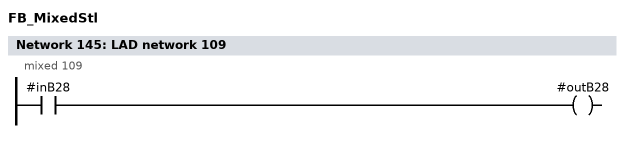
   RUNG wire#powerrail
      Contact( #inB28 )
      Coil( #outB28 )
   END_RUNG
   // the same network as SCL:
   #outB28 := #inB28;
END_REGION

REGION Network 146 (FBD): FBD network 110
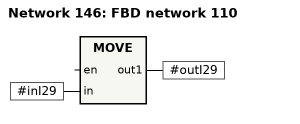
   #outI29 := #inI29;
END_REGION

REGION Network 147 (SCL): SCL network 111
   #tI10 := #inI30 + #cI20;
           IF #inB30 THEN
               #outR10 := #inR10 * 2.0;
           END_IF;
END_REGION

REGION Network 148 (STL): STL network 37
         A     #inB36;
         AN    #stB36;
         =     #outB36;
END_REGION

REGION Network 149: LAD network 112
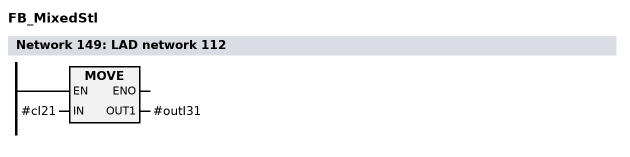
   RUNG wire#powerrail
      Move(in := #cI21, out1 => #outI31)
   END_RUNG
   // the same network as SCL:
   #outI31 := #cI21;
END_REGION

REGION Network 150 (FBD): FBD network 113
   // mixed 113
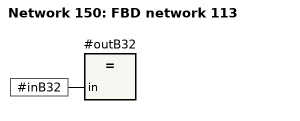
   #outB32 := #inB32;
END_REGION

REGION Network 151 (SCL): SCL network 114
   #tI13 := #inI33 + #cI23;
           IF #inB33 THEN
               #outR13 := #inR13 * 2.0;
           END_IF;
END_REGION

REGION Network 152 (STL): STL network 38
         L     #inI37;
         L     #stI37;
         +I;
         T     #outI37;
END_REGION

REGION Network 153: LAD network 115
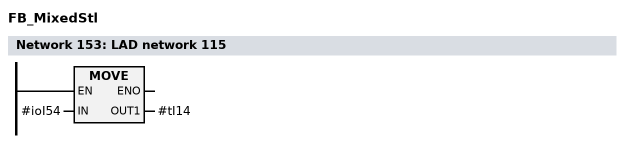
   RUNG wire#powerrail
      Move(in := #ioI54, out1 => #tI14)
   END_RUNG
   // the same network as SCL:
   #tI14 := #ioI54;
END_REGION

REGION Network 154 (FBD): FBD network 116
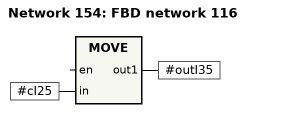
   #outI35 := #cI25;
END_REGION

REGION Network 155 (SCL): SCL network 117
   // mixed 117
   #tI16 := #inI36 + #cI26;
           IF #inB36 THEN
               #outR16 := #inR16 * 2.0;
           END_IF;
END_REGION

REGION Network 156 (STL): STL network 39
         L     #inR18;
         L     #tR38;
         *R;
         T     #outR18;  // product
END_REGION

REGION Network 157: LAD network 118
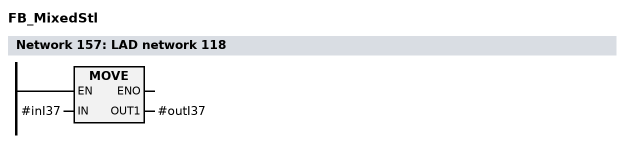
   RUNG wire#powerrail
      Move(in := #inI37, out1 => #outI37)
   END_RUNG
   // the same network as SCL:
   #outI37 := #inI37;
END_REGION

REGION Network 158 (FBD): FBD network 119
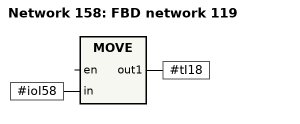
   #tI18 := #ioI58;
END_REGION

REGION Network 159 (SCL): SCL network 120
   #tI19 := #inI39 + #cI29;
           IF #inB39 THEN
               #outR19 := #inR19 * 2.0;
           END_IF;
END_REGION

REGION Network 160 (STL): STL network 40
         A     #inB39;
         AN    #stB39;
         =     #outB39;
END_REGION
END_FUNCTION_BLOCK

FUNCTION "FC_Stl" : Void   // FC1, STL
TITLE = STL test FC
{ S7_Optimized_Access := 'TRUE' }
VERSION : 0.1
   VAR_INPUT
      "a" : Bool;
      "b" : Bool;
      x : Int;
      y : Int;
   END_VAR
   VAR_OUTPUT
      q : Bool;
      sum : Int;
   END_VAR
   VAR_TEMP
      t : Int;
   END_VAR
BEGIN

REGION Network 1: Bit logic
   // Network comment line 1
         A     #"a";  // and a
         AN    #"b";
         =     #q;
END_REGION

REGION Network 2: Arithmetic
         L     #x;
         L     #y;
         +I;
         T     #t;

         L     #t;
         L     0;
         >I;
         JC    M001;
         L     0;
         T     #t;
   M001: L     #t;
         T     #sum;
END_REGION
END_FUNCTION

FUNCTION "FC_StlNoPar" : Void   // FC2, STL
{ S7_Optimized_Access := 'FALSE' }
VERSION : 0.1
BEGIN

REGION Network 1
         NOP   0;
END_REGION
END_FUNCTION

FUNCTION "FC_StlPar" : Void   // FC3, STL
{ S7_Optimized_Access := 'TRUE' }
VERSION : 0.1
   VAR_INPUT
      x : Int;
      y : Int;
   END_VAR
   VAR_OUTPUT
      q : Bool;
      r : Int;
   END_VAR
BEGIN

REGION Network 1
         L     #x;
         L     #y;
         +I;
         T     #r;
         >I;
         =     #q;
END_REGION
END_FUNCTION

FUNCTION "FC_BigFbd" : Void   // FC4, FBD
{ S7_Optimized_Access := 'TRUE' }
VERSION : 0.1
   VAR_INPUT
      inB0 : Bool;   // input bit 0
      inB1 : Bool;
      inB2 : Bool;
      inB3 : Bool;
      inB4 : Bool;
      inB5 : Bool;
      inB6 : Bool;
      inB7 : Bool;
      inB8 : Bool;
      inB9 : Bool;
      inB10 : Bool;   // input bit 10
      inB11 : Bool;
      inB12 : Bool;
      inB13 : Bool;
      inB14 : Bool;
      inB15 : Bool;
      inB16 : Bool;
      inB17 : Bool;
      inB18 : Bool;
      inB19 : Bool;
      inI0 : Int;
      inI1 : Int;
      inI2 : Int;
      inI3 : Int;
      inI4 : Int;
      inI5 : Int;
      inI6 : Int;
      inI7 : Int;
      inI8 : Int;
      inI9 : Int;
      inI10 : Int;
      inI11 : Int;
      inI12 : Int;
      inI13 : Int;
      inI14 : Int;
      inI15 : Int;
      inI16 : Int;
      inI17 : Int;
      inI18 : Int;
      inI19 : Int;
      inR0 : Real;
      inR1 : Real;
      inR2 : Real;
      inR3 : Real;
      inR4 : Real;
      inR5 : Real;
      inR6 : Real;
      inR7 : Real;
      inR8 : Real;
      inR9 : Real;
      inD0 : DInt;
      inD1 : DInt;
      inD2 : DInt;
      inD3 : DInt;
      inD4 : DInt;
      inD5 : DInt;
      inD6 : DInt;
      inD7 : DInt;
      inD8 : DInt;
      inD9 : DInt;
      inArr : Array[0..99] of Int;   // input array
      inStr : String;
      inSt : Struct
         x : Int;
         y : Real;
         z : Bool;
      END_STRUCT;
   END_VAR
   VAR_OUTPUT
      outB0 : Bool;
      outB1 : Bool;
      outB2 : Bool;
      outB3 : Bool;
      outB4 : Bool;
      outB5 : Bool;
      outB6 : Bool;
      outB7 : Bool;
      outB8 : Bool;
      outB9 : Bool;
      outB10 : Bool;
      outB11 : Bool;
      outB12 : Bool;
      outB13 : Bool;
      outB14 : Bool;
      outB15 : Bool;
      outB16 : Bool;
      outB17 : Bool;
      outB18 : Bool;
      outB19 : Bool;
      outI0 : Int;   // output int 0
      outI1 : Int;
      outI2 : Int;
      outI3 : Int;
      outI4 : Int;
      outI5 : Int;
      outI6 : Int;
      outI7 : Int;
      outI8 : Int;
      outI9 : Int;
      outI10 : Int;   // output int 10
      outI11 : Int;
      outI12 : Int;
      outI13 : Int;
      outI14 : Int;
      outI15 : Int;
      outI16 : Int;
      outI17 : Int;
      outI18 : Int;
      outI19 : Int;
      outR0 : Real;
      outR1 : Real;
      outR2 : Real;
      outR3 : Real;
      outR4 : Real;
      outR5 : Real;
      outR6 : Real;
      outR7 : Real;
      outR8 : Real;
      outR9 : Real;
      outD0 : DInt;
      outD1 : DInt;
      outD2 : DInt;
      outD3 : DInt;
      outD4 : DInt;
      outD5 : DInt;
      outD6 : DInt;
      outD7 : DInt;
      outD8 : DInt;
      outD9 : DInt;
   END_VAR
   VAR_IN_OUT
      ioI0 : Int;
      ioI1 : Int;
   END_VAR
   VAR_TEMP
      tI0 : Int;
      tI1 : Int;
      tI2 : Int;
      tI3 : Int;
      tI4 : Int;
      tI5 : Int;
      tI6 : Int;
      tI7 : Int;
      tI8 : Int;
      tI9 : Int;
      tI10 : Int;
      tI11 : Int;
      tI12 : Int;
      tI13 : Int;
      tI14 : Int;
      tI15 : Int;
      tI16 : Int;
      tI17 : Int;
      tI18 : Int;
      tI19 : Int;
      tI20 : Int;
      tI21 : Int;
      tI22 : Int;
      tI23 : Int;
      tI24 : Int;
      tI25 : Int;
      tI26 : Int;
      tI27 : Int;
      tI28 : Int;
      tI29 : Int;
      tI30 : Int;
      tI31 : Int;
      tI32 : Int;
      tI33 : Int;
      tI34 : Int;
      tI35 : Int;
      tI36 : Int;
      tI37 : Int;
      tI38 : Int;
      tI39 : Int;
      tI40 : Int;
      tI41 : Int;
      tI42 : Int;
      tI43 : Int;
      tI44 : Int;
      tI45 : Int;
      tI46 : Int;
      tI47 : Int;
      tI48 : Int;
      tI49 : Int;
      tI50 : Int;
      tI51 : Int;
      tI52 : Int;
      tI53 : Int;
      tI54 : Int;
      tI55 : Int;
      tI56 : Int;
      tI57 : Int;
      tI58 : Int;
      tI59 : Int;
      tI60 : Int;
      tI61 : Int;
      tI62 : Int;
      tI63 : Int;
      tI64 : Int;
      tI65 : Int;
      tI66 : Int;
      tI67 : Int;
      tI68 : Int;
      tI69 : Int;
      tI70 : Int;
      tI71 : Int;
      tI72 : Int;
      tI73 : Int;
      tI74 : Int;
      tI75 : Int;
      tI76 : Int;
      tI77 : Int;
      tI78 : Int;
      tI79 : Int;
      tI80 : Int;
      tI81 : Int;
      tI82 : Int;
      tI83 : Int;
      tI84 : Int;
      tI85 : Int;
      tI86 : Int;
      tI87 : Int;
      tI88 : Int;
      tI89 : Int;
      tI90 : Int;
      tI91 : Int;
      tI92 : Int;
      tI93 : Int;
      tI94 : Int;
      tI95 : Int;
      tI96 : Int;
      tI97 : Int;
      tI98 : Int;
      tI99 : Int;
      tR0 : Real;
      tR1 : Real;
      tR2 : Real;
      tR3 : Real;
      tR4 : Real;
      tR5 : Real;
      tR6 : Real;
      tR7 : Real;
      tR8 : Real;
      tR9 : Real;
      tR10 : Real;
      tR11 : Real;
      tR12 : Real;
      tR13 : Real;
      tR14 : Real;
      tR15 : Real;
      tR16 : Real;
      tR17 : Real;
      tR18 : Real;
      tR19 : Real;
      tR20 : Real;
      tR21 : Real;
      tR22 : Real;
      tR23 : Real;
      tR24 : Real;
      tR25 : Real;
      tR26 : Real;
      tR27 : Real;
      tR28 : Real;
      tR29 : Real;
      tR30 : Real;
      tR31 : Real;
      tR32 : Real;
      tR33 : Real;
      tR34 : Real;
      tR35 : Real;
      tR36 : Real;
      tR37 : Real;
      tR38 : Real;
      tR39 : Real;
      tR40 : Real;
      tR41 : Real;
      tR42 : Real;
      tR43 : Real;
      tR44 : Real;
      tR45 : Real;
      tR46 : Real;
      tR47 : Real;
      tR48 : Real;
      tR49 : Real;
   END_VAR
   VAR CONSTANT
      cI0 : Int := 0;
      cI1 : Int := 3;
      cI2 : Int := 6;
      cI3 : Int := 9;
      cI4 : Int := 12;
      cI5 : Int := 15;
      cI6 : Int := 18;
      cI7 : Int := 21;
      cI8 : Int := 24;
      cI9 : Int := 27;
      cI10 : Int := 30;
      cI11 : Int := 33;
      cI12 : Int := 36;
      cI13 : Int := 39;
      cI14 : Int := 42;
      cI15 : Int := 45;
      cI16 : Int := 48;
      cI17 : Int := 51;
      cI18 : Int := 54;
      cI19 : Int := 57;
      cI20 : Int := 60;
      cI21 : Int := 63;
      cI22 : Int := 66;
      cI23 : Int := 69;
      cI24 : Int := 72;
      cI25 : Int := 75;
      cI26 : Int := 78;
      cI27 : Int := 81;
      cI28 : Int := 84;
      cI29 : Int := 87;
   END_VAR
BEGIN

REGION Network 1: FBD network 1
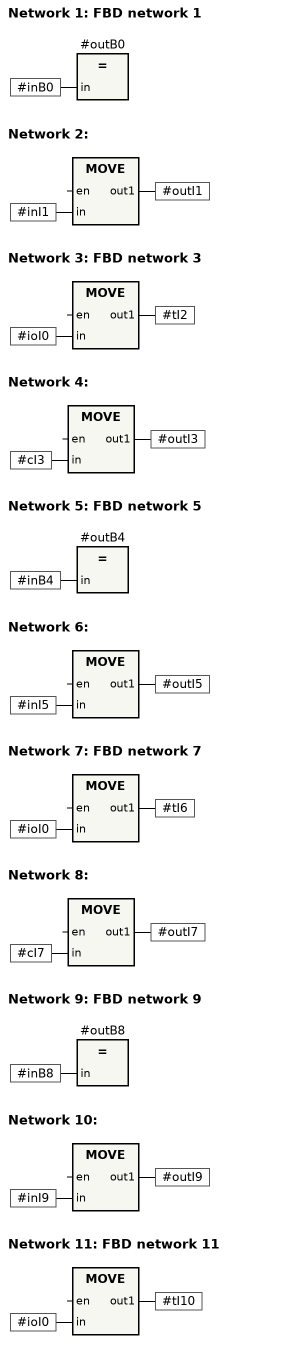
   #outB0 := #inB0;
END_REGION

REGION Network 2
   #outI1 := #inI1;
END_REGION

REGION Network 3: FBD network 3
   #tI2 := #ioI0;
END_REGION

REGION Network 4
   #outI3 := #cI3;
END_REGION

REGION Network 5: FBD network 5
   #outB4 := #inB4;
END_REGION

REGION Network 6
   #outI5 := #inI5;
END_REGION

REGION Network 7: FBD network 7
   #tI6 := #ioI0;
END_REGION

REGION Network 8
   #outI7 := #cI7;
END_REGION

REGION Network 9: FBD network 9
   #outB8 := #inB8;
END_REGION

REGION Network 10
   #outI9 := #inI9;
END_REGION

REGION Network 11: FBD network 11
   #tI10 := #ioI0;
END_REGION

REGION Network 12
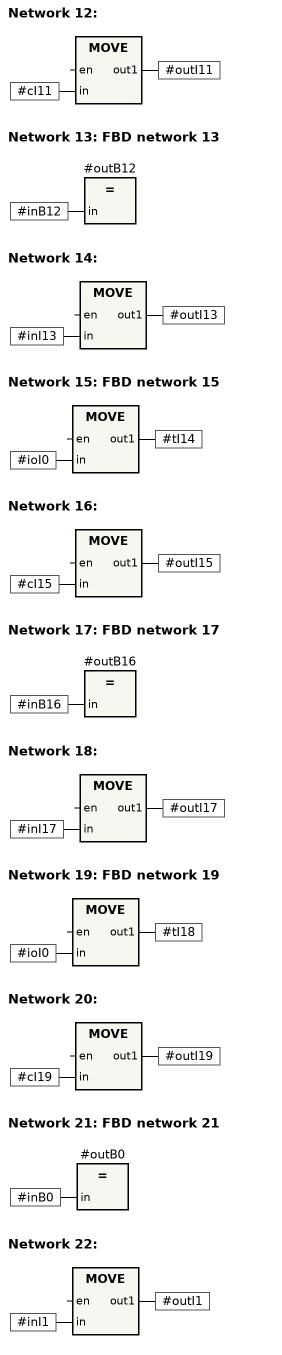
   #outI11 := #cI11;
END_REGION

REGION Network 13: FBD network 13
   #outB12 := #inB12;
END_REGION

REGION Network 14
   #outI13 := #inI13;
END_REGION

REGION Network 15: FBD network 15
   #tI14 := #ioI0;
END_REGION

REGION Network 16
   #outI15 := #cI15;
END_REGION

REGION Network 17: FBD network 17
   #outB16 := #inB16;
END_REGION

REGION Network 18
   #outI17 := #inI17;
END_REGION

REGION Network 19: FBD network 19
   #tI18 := #ioI0;
END_REGION

REGION Network 20
   #outI19 := #cI19;
END_REGION

REGION Network 21: FBD network 21
   #outB0 := #inB0;
END_REGION

REGION Network 22
   #outI1 := #inI1;
END_REGION

REGION Network 23: FBD network 23
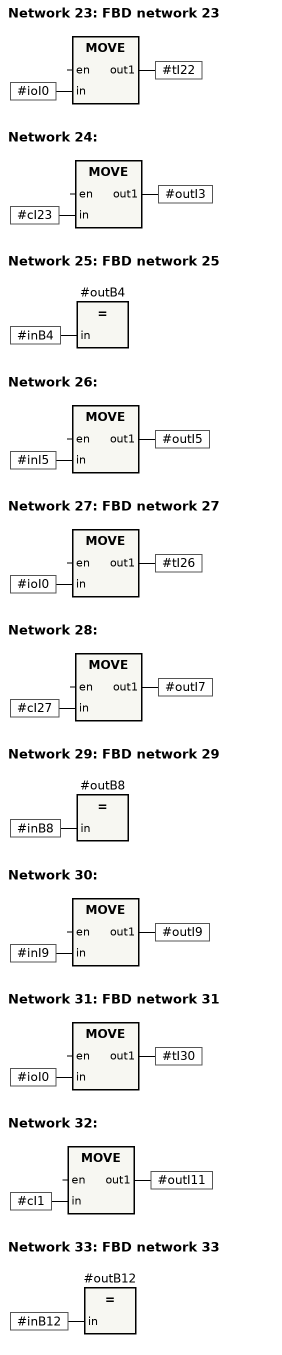
   #tI22 := #ioI0;
END_REGION

REGION Network 24
   #outI3 := #cI23;
END_REGION

REGION Network 25: FBD network 25
   #outB4 := #inB4;
END_REGION

REGION Network 26
   #outI5 := #inI5;
END_REGION

REGION Network 27: FBD network 27
   #tI26 := #ioI0;
END_REGION

REGION Network 28
   #outI7 := #cI27;
END_REGION

REGION Network 29: FBD network 29
   #outB8 := #inB8;
END_REGION

REGION Network 30
   #outI9 := #inI9;
END_REGION

REGION Network 31: FBD network 31
   #tI30 := #ioI0;
END_REGION

REGION Network 32
   #outI11 := #cI1;
END_REGION

REGION Network 33: FBD network 33
   #outB12 := #inB12;
END_REGION

REGION Network 34
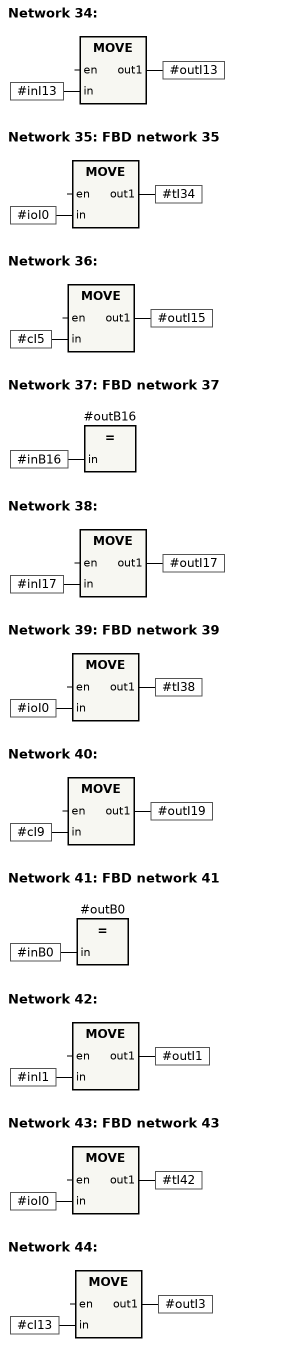
   #outI13 := #inI13;
END_REGION

REGION Network 35: FBD network 35
   #tI34 := #ioI0;
END_REGION

REGION Network 36
   #outI15 := #cI5;
END_REGION

REGION Network 37: FBD network 37
   #outB16 := #inB16;
END_REGION

REGION Network 38
   #outI17 := #inI17;
END_REGION

REGION Network 39: FBD network 39
   #tI38 := #ioI0;
END_REGION

REGION Network 40
   #outI19 := #cI9;
END_REGION

REGION Network 41: FBD network 41
   #outB0 := #inB0;
END_REGION

REGION Network 42
   #outI1 := #inI1;
END_REGION

REGION Network 43: FBD network 43
   #tI42 := #ioI0;
END_REGION

REGION Network 44
   #outI3 := #cI13;
END_REGION

REGION Network 45: FBD network 45
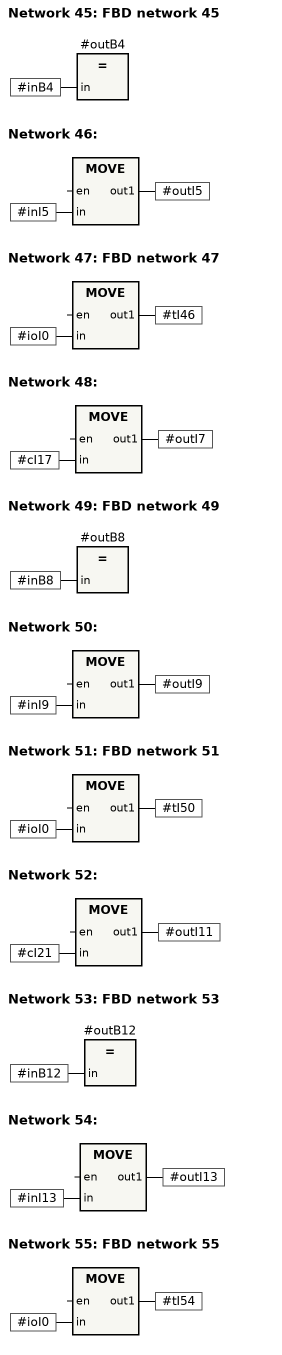
   #outB4 := #inB4;
END_REGION

REGION Network 46
   #outI5 := #inI5;
END_REGION

REGION Network 47: FBD network 47
   #tI46 := #ioI0;
END_REGION

REGION Network 48
   #outI7 := #cI17;
END_REGION

REGION Network 49: FBD network 49
   #outB8 := #inB8;
END_REGION

REGION Network 50
   #outI9 := #inI9;
END_REGION

REGION Network 51: FBD network 51
   #tI50 := #ioI0;
END_REGION

REGION Network 52
   #outI11 := #cI21;
END_REGION

REGION Network 53: FBD network 53
   #outB12 := #inB12;
END_REGION

REGION Network 54
   #outI13 := #inI13;
END_REGION

REGION Network 55: FBD network 55
   #tI54 := #ioI0;
END_REGION

REGION Network 56
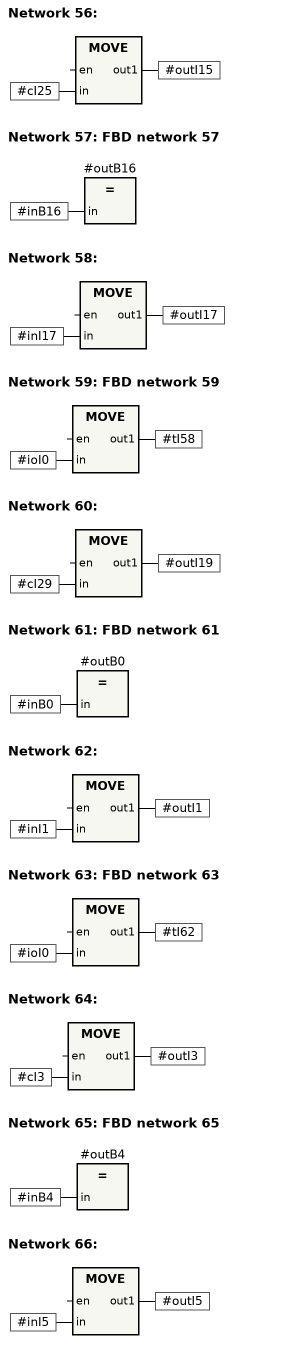
   #outI15 := #cI25;
END_REGION

REGION Network 57: FBD network 57
   #outB16 := #inB16;
END_REGION

REGION Network 58
   #outI17 := #inI17;
END_REGION

REGION Network 59: FBD network 59
   #tI58 := #ioI0;
END_REGION

REGION Network 60
   #outI19 := #cI29;
END_REGION

REGION Network 61: FBD network 61
   #outB0 := #inB0;
END_REGION

REGION Network 62
   #outI1 := #inI1;
END_REGION

REGION Network 63: FBD network 63
   #tI62 := #ioI0;
END_REGION

REGION Network 64
   #outI3 := #cI3;
END_REGION

REGION Network 65: FBD network 65
   #outB4 := #inB4;
END_REGION

REGION Network 66
   #outI5 := #inI5;
END_REGION

REGION Network 67: FBD network 67
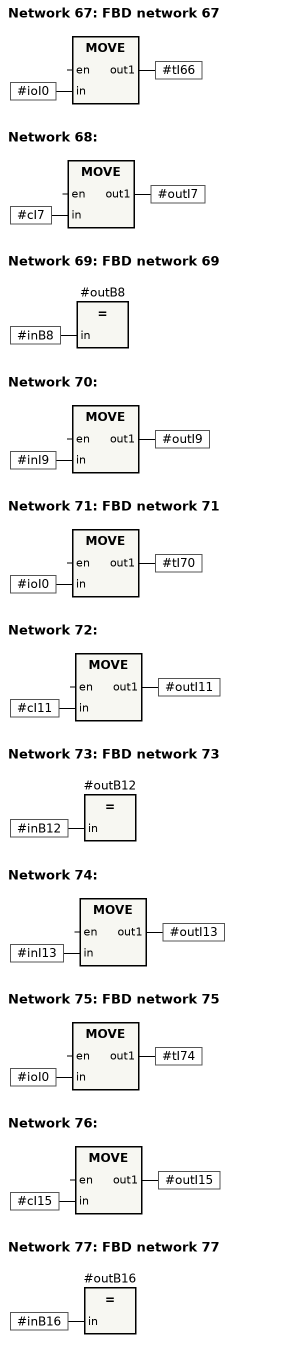
   #tI66 := #ioI0;
END_REGION

REGION Network 68
   #outI7 := #cI7;
END_REGION

REGION Network 69: FBD network 69
   #outB8 := #inB8;
END_REGION

REGION Network 70
   #outI9 := #inI9;
END_REGION

REGION Network 71: FBD network 71
   #tI70 := #ioI0;
END_REGION

REGION Network 72
   #outI11 := #cI11;
END_REGION

REGION Network 73: FBD network 73
   #outB12 := #inB12;
END_REGION

REGION Network 74
   #outI13 := #inI13;
END_REGION

REGION Network 75: FBD network 75
   #tI74 := #ioI0;
END_REGION

REGION Network 76
   #outI15 := #cI15;
END_REGION

REGION Network 77: FBD network 77
   #outB16 := #inB16;
END_REGION

REGION Network 78
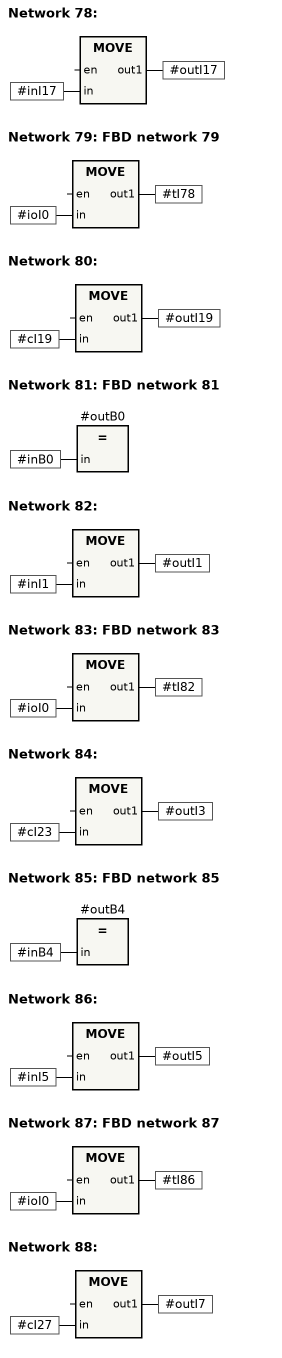
   #outI17 := #inI17;
END_REGION

REGION Network 79: FBD network 79
   #tI78 := #ioI0;
END_REGION

REGION Network 80
   #outI19 := #cI19;
END_REGION

REGION Network 81: FBD network 81
   #outB0 := #inB0;
END_REGION

REGION Network 82
   #outI1 := #inI1;
END_REGION

REGION Network 83: FBD network 83
   #tI82 := #ioI0;
END_REGION

REGION Network 84
   #outI3 := #cI23;
END_REGION

REGION Network 85: FBD network 85
   #outB4 := #inB4;
END_REGION

REGION Network 86
   #outI5 := #inI5;
END_REGION

REGION Network 87: FBD network 87
   #tI86 := #ioI0;
END_REGION

REGION Network 88
   #outI7 := #cI27;
END_REGION

REGION Network 89: FBD network 89
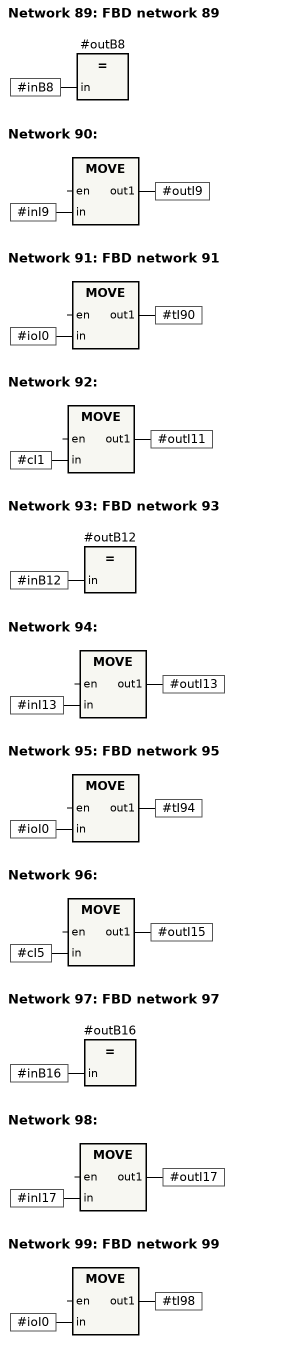
   #outB8 := #inB8;
END_REGION

REGION Network 90
   #outI9 := #inI9;
END_REGION

REGION Network 91: FBD network 91
   #tI90 := #ioI0;
END_REGION

REGION Network 92
   #outI11 := #cI1;
END_REGION

REGION Network 93: FBD network 93
   #outB12 := #inB12;
END_REGION

REGION Network 94
   #outI13 := #inI13;
END_REGION

REGION Network 95: FBD network 95
   #tI94 := #ioI0;
END_REGION

REGION Network 96
   #outI15 := #cI5;
END_REGION

REGION Network 97: FBD network 97
   #outB16 := #inB16;
END_REGION

REGION Network 98
   #outI17 := #inI17;
END_REGION

REGION Network 99: FBD network 99
   #tI98 := #ioI0;
END_REGION

REGION Network 100
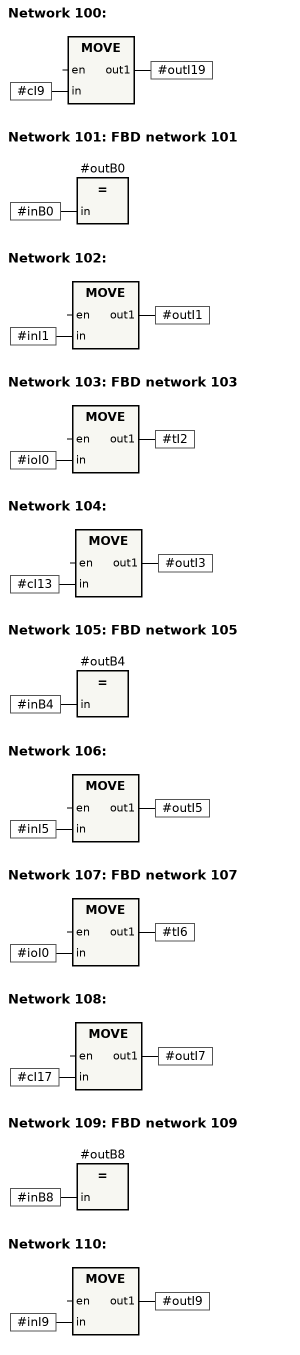
   #outI19 := #cI9;
END_REGION

REGION Network 101: FBD network 101
   #outB0 := #inB0;
END_REGION

REGION Network 102
   #outI1 := #inI1;
END_REGION

REGION Network 103: FBD network 103
   #tI2 := #ioI0;
END_REGION

REGION Network 104
   #outI3 := #cI13;
END_REGION

REGION Network 105: FBD network 105
   #outB4 := #inB4;
END_REGION

REGION Network 106
   #outI5 := #inI5;
END_REGION

REGION Network 107: FBD network 107
   #tI6 := #ioI0;
END_REGION

REGION Network 108
   #outI7 := #cI17;
END_REGION

REGION Network 109: FBD network 109
   #outB8 := #inB8;
END_REGION

REGION Network 110
   #outI9 := #inI9;
END_REGION

REGION Network 111: FBD network 111
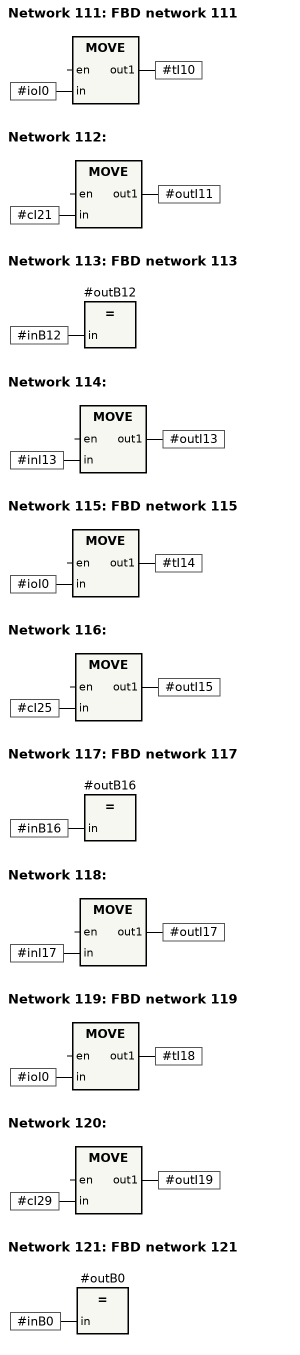
   #tI10 := #ioI0;
END_REGION

REGION Network 112
   #outI11 := #cI21;
END_REGION

REGION Network 113: FBD network 113
   #outB12 := #inB12;
END_REGION

REGION Network 114
   #outI13 := #inI13;
END_REGION

REGION Network 115: FBD network 115
   #tI14 := #ioI0;
END_REGION

REGION Network 116
   #outI15 := #cI25;
END_REGION

REGION Network 117: FBD network 117
   #outB16 := #inB16;
END_REGION

REGION Network 118
   #outI17 := #inI17;
END_REGION

REGION Network 119: FBD network 119
   #tI18 := #ioI0;
END_REGION

REGION Network 120
   #outI19 := #cI29;
END_REGION

REGION Network 121: FBD network 121
   #outB0 := #inB0;
END_REGION

REGION Network 122
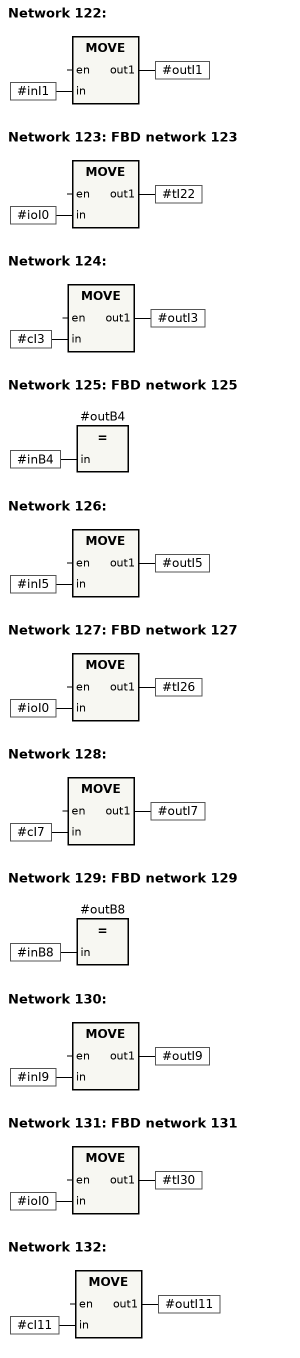
   #outI1 := #inI1;
END_REGION

REGION Network 123: FBD network 123
   #tI22 := #ioI0;
END_REGION

REGION Network 124
   #outI3 := #cI3;
END_REGION

REGION Network 125: FBD network 125
   #outB4 := #inB4;
END_REGION

REGION Network 126
   #outI5 := #inI5;
END_REGION

REGION Network 127: FBD network 127
   #tI26 := #ioI0;
END_REGION

REGION Network 128
   #outI7 := #cI7;
END_REGION

REGION Network 129: FBD network 129
   #outB8 := #inB8;
END_REGION

REGION Network 130
   #outI9 := #inI9;
END_REGION

REGION Network 131: FBD network 131
   #tI30 := #ioI0;
END_REGION

REGION Network 132
   #outI11 := #cI11;
END_REGION

REGION Network 133: FBD network 133
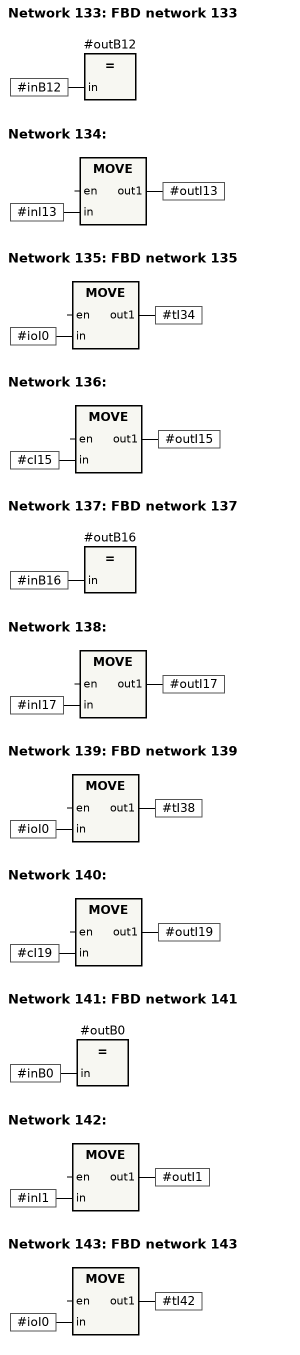
   #outB12 := #inB12;
END_REGION

REGION Network 134
   #outI13 := #inI13;
END_REGION

REGION Network 135: FBD network 135
   #tI34 := #ioI0;
END_REGION

REGION Network 136
   #outI15 := #cI15;
END_REGION

REGION Network 137: FBD network 137
   #outB16 := #inB16;
END_REGION

REGION Network 138
   #outI17 := #inI17;
END_REGION

REGION Network 139: FBD network 139
   #tI38 := #ioI0;
END_REGION

REGION Network 140
   #outI19 := #cI19;
END_REGION

REGION Network 141: FBD network 141
   #outB0 := #inB0;
END_REGION

REGION Network 142
   #outI1 := #inI1;
END_REGION

REGION Network 143: FBD network 143
   #tI42 := #ioI0;
END_REGION

REGION Network 144
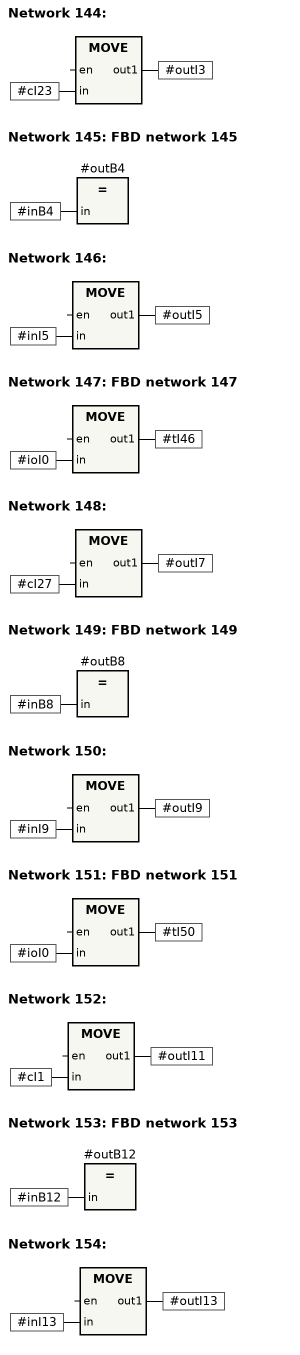
   #outI3 := #cI23;
END_REGION

REGION Network 145: FBD network 145
   #outB4 := #inB4;
END_REGION

REGION Network 146
   #outI5 := #inI5;
END_REGION

REGION Network 147: FBD network 147
   #tI46 := #ioI0;
END_REGION

REGION Network 148
   #outI7 := #cI27;
END_REGION

REGION Network 149: FBD network 149
   #outB8 := #inB8;
END_REGION

REGION Network 150
   #outI9 := #inI9;
END_REGION

REGION Network 151: FBD network 151
   #tI50 := #ioI0;
END_REGION

REGION Network 152
   #outI11 := #cI1;
END_REGION

REGION Network 153: FBD network 153
   #outB12 := #inB12;
END_REGION

REGION Network 154
   #outI13 := #inI13;
END_REGION

REGION Network 155: FBD network 155
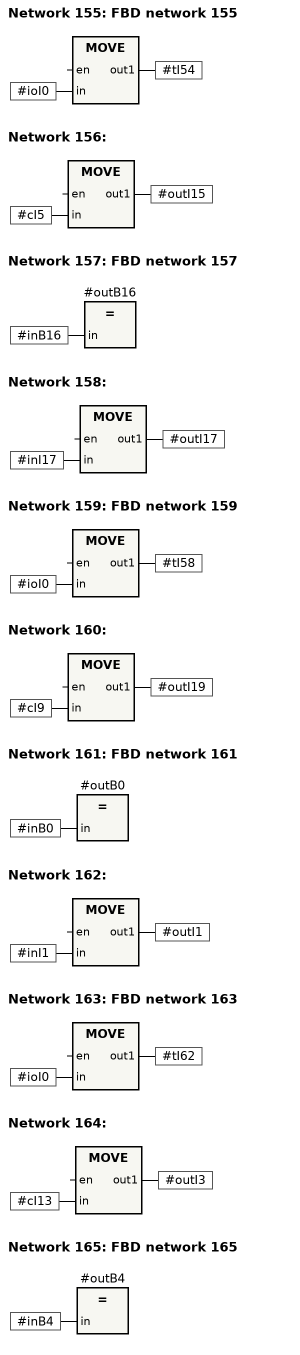
   #tI54 := #ioI0;
END_REGION

REGION Network 156
   #outI15 := #cI5;
END_REGION

REGION Network 157: FBD network 157
   #outB16 := #inB16;
END_REGION

REGION Network 158
   #outI17 := #inI17;
END_REGION

REGION Network 159: FBD network 159
   #tI58 := #ioI0;
END_REGION

REGION Network 160
   #outI19 := #cI9;
END_REGION

REGION Network 161: FBD network 161
   #outB0 := #inB0;
END_REGION

REGION Network 162
   #outI1 := #inI1;
END_REGION

REGION Network 163: FBD network 163
   #tI62 := #ioI0;
END_REGION

REGION Network 164
   #outI3 := #cI13;
END_REGION

REGION Network 165: FBD network 165
   #outB4 := #inB4;
END_REGION

REGION Network 166
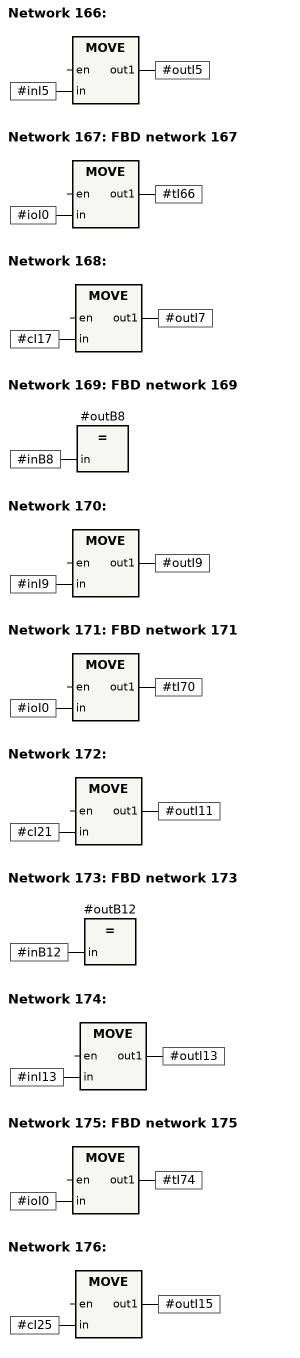
   #outI5 := #inI5;
END_REGION

REGION Network 167: FBD network 167
   #tI66 := #ioI0;
END_REGION

REGION Network 168
   #outI7 := #cI17;
END_REGION

REGION Network 169: FBD network 169
   #outB8 := #inB8;
END_REGION

REGION Network 170
   #outI9 := #inI9;
END_REGION

REGION Network 171: FBD network 171
   #tI70 := #ioI0;
END_REGION

REGION Network 172
   #outI11 := #cI21;
END_REGION

REGION Network 173: FBD network 173
   #outB12 := #inB12;
END_REGION

REGION Network 174
   #outI13 := #inI13;
END_REGION

REGION Network 175: FBD network 175
   #tI74 := #ioI0;
END_REGION

REGION Network 176
   #outI15 := #cI25;
END_REGION

REGION Network 177: FBD network 177
